Fanuc KAREL source: KO00058.KL

PROGRAM KO00058
%NOLOCKGROUP
%ENVIRONMENT MIR
VAR
  P1: XYZWPR
  P2: XYZWPREXT
  F: BOOLEAN
  OUT: XYZWPR
BEGIN
  F = TRUE
  OUT = MIRROR(P1, P2, F)
END KO00058
